FUNCTION_BLOCK FB_EventLoggerListener EXTENDS FB_ListenerBase2
VAR_INPUT
END_VAR
VAR_OUTPUT
END_VAR
VAR
	sJsonAttribute : STRING (10000);	
	hr : HRESULT;
	
	nCntMessagesSent : INT;
	nCntAlarmsRaised : INT;
	nCntAlarmsConfirmed : INT;
	nCntAlarmsCleared : INT;
	
	//text retrieval of message
	fbRequestEventText : FB_RequestEventText;
	{attribute 'TcEncoding':='UTF-8'}
	sLastMessageText : STRING;
	bReqText : BOOL;
	
	aAlarmHistory : ARRAY[1..MAX_ALARMS_HISTORY] OF ST_AlarmHistoryEntry;
    i : INT;
    
    // Zmienne tymczasowe, czekające na pobranie tekstu
    nTempTimestamp : ULINT;
    eTempSeverity  : TcEventSeverity;
END_VAR
VAR CONSTANT
    MAX_ALARMS_HISTORY : INT := 20; // Rozmiar tablicy (np. 20 ostatnich alarmów)
END_VAR

METHOD Execute : HRESULT
VAR_INPUT
END_VAR
Execute := SUPER^.Execute(); //retrieve events

// Zmodyfikowany kod odbioru tekstu
IF bReqText AND NOT fbRequestEventText.bBusy THEN
    
    // 1. Odbierz tekst lub ustaw błąd
    IF fbRequestEventText.bError THEN 
        sLastMessageText := 'Error retrieving text';
    ELSE
        fbRequestEventText.GetString(sLastMessageText, SIZEOF(sLastMessageText));
    END_IF
    
    bReqText := FALSE; 
    
    // 2. Przesuń starsze alarmy w tablicy (zwolnij indeks 1)
    FOR i := MAX_ALARMS_HISTORY TO 2 BY -1 DO
        aAlarmHistory[i] := aAlarmHistory[i-1];
    END_FOR
    
    // 3. Wpisz najnowszy alarm na indeks 1
    aAlarmHistory[1].sMessageText := sLastMessageText;
    aAlarmHistory[1].nTimestamp   := nTempTimestamp;
    aAlarmHistory[1].eSeverity    := eTempSeverity;

END_IF
END_METHOD

METHOD OnAlarmCleared : HRESULT
VAR_INPUT
	fbEvent : REFERENCE TO FB_TcEvent;
END_VAR
nCntAlarmsCleared := nCntAlarmsCleared + 1;

OnAlarmCleared := S_OK; // in order to receive more callbacks (Set <> S_OK in order to cancel the callbacks for this program cycle.)
END_METHOD

METHOD OnAlarmConfirmed : HRESULT
VAR_INPUT
	fbEvent : REFERENCE TO FB_TcEvent;
END_VAR
nCntAlarmsConfirmed := nCntAlarmsConfirmed + 1;

OnAlarmConfirmed := S_OK; // in order to receive more callbacks (Set <> S_OK in order to cancel the callbacks for this program cycle.)
END_METHOD

METHOD OnAlarmRaised : HRESULT
VAR_INPUT
    fbEvent : REFERENCE TO FB_TcEvent;
END_VAR


// Wewnątrz metody:
hr := fbEvent.GetJsonAttribute(sJsonAttribute, SIZEOF(sJsonAttribute));
nCntAlarmsRaised := nCntAlarmsRaised + 1;

// --- ZAPISZ DANE DO ZMIENNYCH TYMCZASOWYCH ---
nTempTimestamp := fbEvent.nTimestamp;
eTempSeverity  := fbEvent.eSeverity;

OnAlarmRaised := S_OK; 
fbRequestEventText.Request(eventClass := fbEvent.EventClass, nEventId := fbEvent.nEventId,
                           nLangId := TcLcid.en_US, ipArgs := fbEvent.ipArguments);
bReqText := TRUE;
END_METHOD

METHOD OnMessageSent : HRESULT
VAR_INPUT
	fbEvent : REFERENCE TO FB_TcEvent;
END_VAR

VAR 
END_VAR
hr := fbEvent.GetJsonAttribute(sJsonAttribute, SIZEOF(sJsonAttribute));
nCntMessagesSent := nCntMessagesSent + 1;

nTempTimestamp := fbEvent.nTimestamp;
eTempSeverity  := fbEvent.eSeverity;

fbRequestEventText.Request(eventClass:=fbEvent.EventClass, nEventId:=fbEvent.nEventId, nLangId:=TcLcid.en_US, ipArgs:=fbEvent.ipArguments );
bReqText := TRUE;

OnMessageSent := S_OK; // in order to receive more callbacks (Set <> S_OK in order to cancel the callbacks for this program cycle.)
END_METHOD

END_FUNCTION_BLOCK

(* stored: Version 1.1.0.1, ProductVersion 3.1.4024.15
   POU FB_EventLoggerListener: Id {50ed088d-9a7d-4c16-86a9-e90b487e4982}, SpecialFunc None
   Method Execute: Id {3c7f655d-2c73-41dc-b085-26c5a3b1cef1}
   Method OnAlarmCleared: Id {036602cd-44fc-40d2-99e6-e6b033452290}
   Method OnAlarmConfirmed: Id {efe870ed-8bbd-4c42-9405-bf33d81f12d4}
   Method OnAlarmRaised: Id {1df5b803-888d-4d2d-ab12-93687f9c1a1e}
   Method OnMessageSent: Id {b4dac56d-cfe9-4434-ae5b-afa117054bdb} *)
